TYPE ST_Component :
STRUCT
	sDescription		: STRING;
	rCompWeightFor100L	: REAL;
	
	rMaxPressure		: REAL;
	rMaxTemp			: REAL;
	rMinFlowRate		: REAL;
	
	
	///Val for actual work
	rCompActWeight		: REAL;
	rFlowTarget			: REAL;
	rRpmTarget			: REAL;
	iMixingTime			: UINT;
	
	//Ctrl
	iLocationInList		: USINT;
	bCtrlByFlowRate		: BOOL;
	bComponentEnable	: BOOL;
	bIsWater			: BOOL;
END_STRUCT
END_TYPE

(* stored: Version 1.1.0.1, ProductVersion 3.1.4024.12
   DUT ST_Component: Id {1e51c929-826d-4c0f-8f5b-13bba334a463} *)
